TYPE ST_MB_WriteRegs :
STRUCT
END_STRUCT
END_TYPE

(* stored: Version 1.1.0.1, ProductVersion 3.1.4024.13
   DUT ST_MB_WriteRegs: Id {2af35b66-be41-46e8-8f04-76528ce150d2} *)
